TYPE ST_BECKHOFFDRIVE_REF : FB_BECKHOFFDRIVE_REF;
END_TYPE

(* stored: Version 1.1.0.1, ProductVersion 3.1.4024.15
   DUT ST_BECKHOFFDRIVE_REF: Id {cbc143a1-5ac6-418f-9b18-417f94979db0} *)
